Fanuc KAREL source: KO00096.KL

PROGRAM KO00096
%NOLOCKGROUP
%ENVIRONMENT MIR
VAR
  P1: JOINTPOS
  P2: JOINTPOS
  F: BOOLEAN
  OUT: JOINTPOS
BEGIN
  F = TRUE
  OUT = MIRROR(P1, P2, F)
END KO00096
